// TIA Portal V21 export
// export: Created 2026-11-22T02:34:48.5366465Z, ExportSetting WithDefaults, DisplayName Totally Integrated Automation Portal, DisplayVersion V21 Update 3, DisplayName STEP 7 Professional, DisplayVersion V21 Update 3, DisplayName STEP 7 Safety, DisplayVersion V21, DisplayName Tech WebApplication, DisplayVersion V21, DisplayName WinCC Basic/Comfort/Advanced, DisplayVersion V21 Update 3, DisplayName WinCC Unified, DisplayVersion V21 Update 3
VBScript "SetS1"  Type=Sub
  SmartTags("D_State") = 1
  SmartTags("D_Bool") = False
  SmartTags("D_SInt") = -128
  SmartTags("D_Int") = -32768
  SmartTags("D_DInt") = -2147483648
  SmartTags("D_USInt") = 0
  SmartTags("D_UInt") = 0
  SmartTags("D_UDInt") = 0
  SmartTags("D_Real") = -999.999
  SmartTags("D_LReal") = -0.00000015
  SmartTags("D_String") = ""
  SmartTags("D_DateTime") = DateSerial(1990, 1, 1) + TimeSerial(0, 0, 0)
  SmartTags("D_Pct") = 0
  SmartTags("D_Range") = 5
  SmartTags("D_Bits") = 1
  SmartTags("D_Vis") = False
  SmartTags("D_En") = False
  SmartTags("D_X") = 10
  SmartTags("D_Y") = 10
  SmartTags("D_Max") = 100
  SmartTags("D_Min") = 0
  SmartTags("D_TL") = -5
  SmartTags("D_BarR") = -5
